{attribute 'qualified_only'}
{attribute 'strict'}
{attribute 'to_string'}
TYPE E_BytesEncoding :
(
	hex := 0,
	base64
);
END_TYPE

(* stored: Version 1.1.0.1
   EnumerationTextList E_BytesEncoding: Id {d960b8fb-3c23-44de-b8b9-be57b73a81aa} *)
